Yaskawa INFORM job: KANT1.JBI

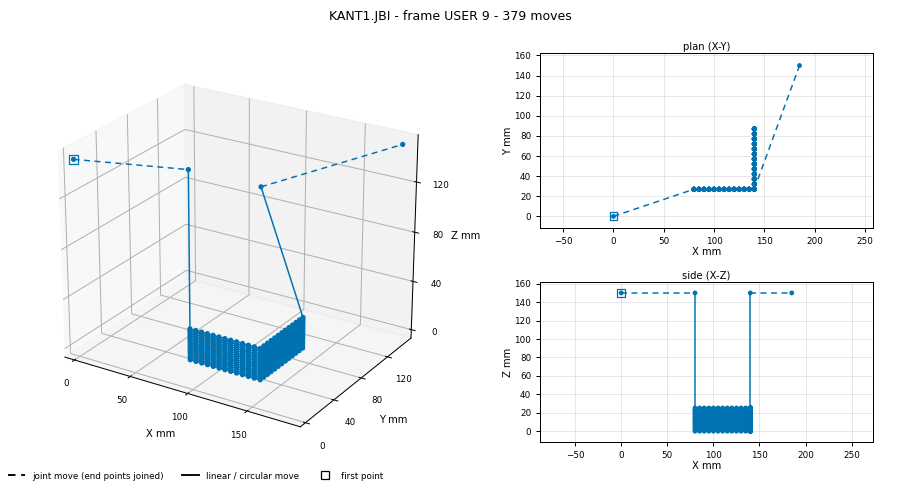
[picture p0: tool path of KANT1.JBI in frame USER 9, 379 of 379 moves have a stored position in this frame; points joined in program order, loops and branches not executed]
/JOB
//NAME KANT1
//POS
///NPOS 379,0,0,0,0,0
///USER 9
///TOOL 1
///POSTYPE USER
///RECTAN
///RCONF 1,0,0,0,0,0,0,0,0,0,0,0,0,0,0,0,0,0,0,0,0,0,0,0
C00000=0.000,0.000,150.000,0.0000,0.0000,-170.0000
C00001=80.000,27.000,150.000,0.0000,0.0000,-170.0000
C00002=80.000,27.000,0.000,0.0000,0.0000,-170.0000
C00003=85.000,27.000,0.000,0.0000,0.0000,-170.0000
C00004=90.000,27.000,0.000,0.0000,0.0000,-170.0000
C00005=95.000,27.000,0.000,0.0000,0.0000,-170.0000
C00006=100.000,27.000,0.000,0.0000,0.0000,-170.0000
C00007=105.000,27.000,0.000,0.0000,0.0000,-170.0000
C00008=110.000,27.000,0.000,0.0000,0.0000,-170.0000
C00009=115.000,27.000,0.000,0.0000,0.0000,-170.0000
C00010=120.000,27.000,0.000,0.0000,0.0000,-170.0000
C00011=125.000,27.000,0.000,0.0000,0.0000,-170.0000
C00012=130.000,27.000,0.000,0.0000,0.0000,-170.0000
C00013=135.000,27.000,0.000,0.0000,0.0000,-170.0000
C00014=140.000,27.000,0.000,0.0000,0.0000,-170.0000
C00015=140.000,32.000,0.000,0.0000,0.0000,-170.0000
C00016=140.000,37.000,0.000,0.0000,0.0000,-170.0000
C00017=140.000,42.000,0.000,0.0000,0.0000,-170.0000
C00018=140.000,47.000,0.000,0.0000,0.0000,-170.0000
C00019=140.000,52.000,0.000,0.0000,0.0000,-170.0000
C00020=140.000,57.000,0.000,0.0000,0.0000,-170.0000
C00021=140.000,62.000,0.000,0.0000,0.0000,-170.0000
C00022=140.000,67.000,0.000,0.0000,0.0000,-170.0000
C00023=140.000,72.000,0.000,0.0000,0.0000,-170.0000
C00024=140.000,77.000,0.000,0.0000,0.0000,-170.0000
C00025=140.000,82.000,0.000,0.0000,0.0000,-170.0000
C00026=140.000,87.000,0.000,0.0000,0.0000,-170.0000
C00027=140.000,87.000,1.800,0.0000,0.0000,-170.0000
C00028=140.000,82.000,1.800,0.0000,0.0000,-170.0000
C00029=140.000,77.000,1.800,0.0000,0.0000,-170.0000
C00030=140.000,72.000,1.800,0.0000,0.0000,-170.0000
C00031=140.000,67.000,1.800,0.0000,0.0000,-170.0000
C00032=140.000,62.000,1.800,0.0000,0.0000,-170.0000
C00033=140.000,57.000,1.800,0.0000,0.0000,-170.0000
C00034=140.000,52.000,1.800,0.0000,0.0000,-170.0000
C00035=140.000,47.000,1.800,0.0000,0.0000,-170.0000
C00036=140.000,42.000,1.800,0.0000,0.0000,-170.0000
C00037=140.000,37.000,1.800,0.0000,0.0000,-170.0000
C00038=140.000,32.000,1.800,0.0000,0.0000,-170.0000
C00039=140.000,27.000,1.800,0.0000,0.0000,-170.0000
C00040=135.000,27.000,1.800,0.0000,0.0000,-170.0000
C00041=130.000,27.000,1.800,0.0000,0.0000,-170.0000
C00042=125.000,27.000,1.800,0.0000,0.0000,-170.0000
C00043=120.000,27.000,1.800,0.0000,0.0000,-170.0000
C00044=115.000,27.000,1.800,0.0000,0.0000,-170.0000
C00045=110.000,27.000,1.800,0.0000,0.0000,-170.0000
C00046=105.000,27.000,1.800,0.0000,0.0000,-170.0000
C00047=100.000,27.000,1.800,0.0000,0.0000,-170.0000
C00048=95.000,27.000,1.800,0.0000,0.0000,-170.0000
C00049=90.000,27.000,1.800,0.0000,0.0000,-170.0000
C00050=85.000,27.000,1.800,0.0000,0.0000,-170.0000
C00051=80.000,27.000,1.800,0.0000,0.0000,-170.0000
C00052=80.000,27.000,3.600,0.0000,0.0000,-170.0000
C00053=85.000,27.000,3.600,0.0000,0.0000,-170.0000
C00054=90.000,27.000,3.600,0.0000,0.0000,-170.0000
C00055=95.000,27.000,3.600,0.0000,0.0000,-170.0000
C00056=100.000,27.000,3.600,0.0000,0.0000,-170.0000
C00057=105.000,27.000,3.600,0.0000,0.0000,-170.0000
C00058=110.000,27.000,3.600,0.0000,0.0000,-170.0000
C00059=115.000,27.000,3.600,0.0000,0.0000,-170.0000
C00060=120.000,27.000,3.600,0.0000,0.0000,-170.0000
C00061=125.000,27.000,3.600,0.0000,0.0000,-170.0000
C00062=130.000,27.000,3.600,0.0000,0.0000,-170.0000
C00063=135.000,27.000,3.600,0.0000,0.0000,-170.0000
C00064=140.000,27.000,3.600,0.0000,0.0000,-170.0000
C00065=140.000,32.000,3.600,0.0000,0.0000,-170.0000
C00066=140.000,37.000,3.600,0.0000,0.0000,-170.0000
C00067=140.000,42.000,3.600,0.0000,0.0000,-170.0000
C00068=140.000,47.000,3.600,0.0000,0.0000,-170.0000
C00069=140.000,52.000,3.600,0.0000,0.0000,-170.0000
C00070=140.000,57.000,3.600,0.0000,0.0000,-170.0000
C00071=140.000,62.000,3.600,0.0000,0.0000,-170.0000
C00072=140.000,67.000,3.600,0.0000,0.0000,-170.0000
C00073=140.000,72.000,3.600,0.0000,0.0000,-170.0000
C00074=140.000,77.000,3.600,0.0000,0.0000,-170.0000
C00075=140.000,82.000,3.600,0.0000,0.0000,-170.0000
C00076=140.000,87.000,3.600,0.0000,0.0000,-170.0000
C00077=140.000,87.000,5.400,0.0000,0.0000,-170.0000
C00078=140.000,82.000,5.400,0.0000,0.0000,-170.0000
C00079=140.000,77.000,5.400,0.0000,0.0000,-170.0000
C00080=140.000,72.000,5.400,0.0000,0.0000,-170.0000
C00081=140.000,67.000,5.400,0.0000,0.0000,-170.0000
C00082=140.000,62.000,5.400,0.0000,0.0000,-170.0000
C00083=140.000,57.000,5.400,0.0000,0.0000,-170.0000
C00084=140.000,52.000,5.400,0.0000,0.0000,-170.0000
C00085=140.000,47.000,5.400,0.0000,0.0000,-170.0000
C00086=140.000,42.000,5.400,0.0000,0.0000,-170.0000
C00087=140.000,37.000,5.400,0.0000,0.0000,-170.0000
C00088=140.000,32.000,5.400,0.0000,0.0000,-170.0000
C00089=140.000,27.000,5.400,0.0000,0.0000,-170.0000
C00090=135.000,27.000,5.400,0.0000,0.0000,-170.0000
C00091=130.000,27.000,5.400,0.0000,0.0000,-170.0000
C00092=125.000,27.000,5.400,0.0000,0.0000,-170.0000
C00093=120.000,27.000,5.400,0.0000,0.0000,-170.0000
C00094=115.000,27.000,5.400,0.0000,0.0000,-170.0000
C00095=110.000,27.000,5.400,0.0000,0.0000,-170.0000
C00096=105.000,27.000,5.400,0.0000,0.0000,-170.0000
C00097=100.000,27.000,5.400,0.0000,0.0000,-170.0000
C00098=95.000,27.000,5.400,0.0000,0.0000,-170.0000
C00099=90.000,27.000,5.400,0.0000,0.0000,-170.0000
C00100=85.000,27.000,5.400,0.0000,0.0000,-170.0000
C00101=80.000,27.000,5.400,0.0000,0.0000,-170.0000
C00102=80.000,27.000,7.200,0.0000,0.0000,-170.0000
C00103=85.000,27.000,7.200,0.0000,0.0000,-170.0000
C00104=90.000,27.000,7.200,0.0000,0.0000,-170.0000
C00105=95.000,27.000,7.200,0.0000,0.0000,-170.0000
C00106=100.000,27.000,7.200,0.0000,0.0000,-170.0000
C00107=105.000,27.000,7.200,0.0000,0.0000,-170.0000
C00108=110.000,27.000,7.200,0.0000,0.0000,-170.0000
C00109=115.000,27.000,7.200,0.0000,0.0000,-170.0000
C00110=120.000,27.000,7.200,0.0000,0.0000,-170.0000
C00111=125.000,27.000,7.200,0.0000,0.0000,-170.0000
C00112=130.000,27.000,7.200,0.0000,0.0000,-170.0000
C00113=135.000,27.000,7.200,0.0000,0.0000,-170.0000
C00114=140.000,27.000,7.200,0.0000,0.0000,-170.0000
C00115=140.000,32.000,7.200,0.0000,0.0000,-170.0000
C00116=140.000,37.000,7.200,0.0000,0.0000,-170.0000
C00117=140.000,42.000,7.200,0.0000,0.0000,-170.0000
C00118=140.000,47.000,7.200,0.0000,0.0000,-170.0000
C00119=140.000,52.000,7.200,0.0000,0.0000,-170.0000
C00120=140.000,57.000,7.200,0.0000,0.0000,-170.0000
C00121=140.000,62.000,7.200,0.0000,0.0000,-170.0000
C00122=140.000,67.000,7.200,0.0000,0.0000,-170.0000
C00123=140.000,72.000,7.200,0.0000,0.0000,-170.0000
C00124=140.000,77.000,7.200,0.0000,0.0000,-170.0000
C00125=140.000,82.000,7.200,0.0000,0.0000,-170.0000
C00126=140.000,87.000,7.200,0.0000,0.0000,-170.0000
C00127=140.000,87.000,9.000,0.0000,0.0000,-170.0000
C00128=140.000,82.000,9.000,0.0000,0.0000,-170.0000
C00129=140.000,77.000,9.000,0.0000,0.0000,-170.0000
C00130=140.000,72.000,9.000,0.0000,0.0000,-170.0000
C00131=140.000,67.000,9.000,0.0000,0.0000,-170.0000
C00132=140.000,62.000,9.000,0.0000,0.0000,-170.0000
C00133=140.000,57.000,9.000,0.0000,0.0000,-170.0000
C00134=140.000,52.000,9.000,0.0000,0.0000,-170.0000
C00135=140.000,47.000,9.000,0.0000,0.0000,-170.0000
C00136=140.000,42.000,9.000,0.0000,0.0000,-170.0000
C00137=140.000,37.000,9.000,0.0000,0.0000,-170.0000
C00138=140.000,32.000,9.000,0.0000,0.0000,-170.0000
C00139=140.000,27.000,9.000,0.0000,0.0000,-170.0000
C00140=135.000,27.000,9.000,0.0000,0.0000,-170.0000
C00141=130.000,27.000,9.000,0.0000,0.0000,-170.0000
C00142=125.000,27.000,9.000,0.0000,0.0000,-170.0000
C00143=120.000,27.000,9.000,0.0000,0.0000,-170.0000
C00144=115.000,27.000,9.000,0.0000,0.0000,-170.0000
C00145=110.000,27.000,9.000,0.0000,0.0000,-170.0000
C00146=105.000,27.000,9.000,0.0000,0.0000,-170.0000
C00147=100.000,27.000,9.000,0.0000,0.0000,-170.0000
C00148=95.000,27.000,9.000,0.0000,0.0000,-170.0000
C00149=90.000,27.000,9.000,0.0000,0.0000,-170.0000
C00150=85.000,27.000,9.000,0.0000,0.0000,-170.0000
C00151=80.000,27.000,9.000,0.0000,0.0000,-170.0000
C00152=80.000,27.000,10.800,0.0000,0.0000,-170.0000
C00153=85.000,27.000,10.800,0.0000,0.0000,-170.0000
C00154=90.000,27.000,10.800,0.0000,0.0000,-170.0000
C00155=95.000,27.000,10.800,0.0000,0.0000,-170.0000
C00156=100.000,27.000,10.800,0.0000,0.0000,-170.0000
C00157=105.000,27.000,10.800,0.0000,0.0000,-170.0000
C00158=110.000,27.000,10.800,0.0000,0.0000,-170.0000
C00159=115.000,27.000,10.800,0.0000,0.0000,-170.0000
C00160=120.000,27.000,10.800,0.0000,0.0000,-170.0000
C00161=125.000,27.000,10.800,0.0000,0.0000,-170.0000
C00162=130.000,27.000,10.800,0.0000,0.0000,-170.0000
C00163=135.000,27.000,10.800,0.0000,0.0000,-170.0000
C00164=140.000,27.000,10.800,0.0000,0.0000,-170.0000
C00165=140.000,32.000,10.800,0.0000,0.0000,-170.0000
C00166=140.000,37.000,10.800,0.0000,0.0000,-170.0000
C00167=140.000,42.000,10.800,0.0000,0.0000,-170.0000
C00168=140.000,47.000,10.800,0.0000,0.0000,-170.0000
C00169=140.000,52.000,10.800,0.0000,0.0000,-170.0000
C00170=140.000,57.000,10.800,0.0000,0.0000,-170.0000
C00171=140.000,62.000,10.800,0.0000,0.0000,-170.0000
C00172=140.000,67.000,10.800,0.0000,0.0000,-170.0000
C00173=140.000,72.000,10.800,0.0000,0.0000,-170.0000
C00174=140.000,77.000,10.800,0.0000,0.0000,-170.0000
C00175=140.000,82.000,10.800,0.0000,0.0000,-170.0000
C00176=140.000,87.000,10.800,0.0000,0.0000,-170.0000
C00177=140.000,87.000,12.600,0.0000,0.0000,-170.0000
C00178=140.000,82.000,12.600,0.0000,0.0000,-170.0000
C00179=140.000,77.000,12.600,0.0000,0.0000,-170.0000
C00180=140.000,72.000,12.600,0.0000,0.0000,-170.0000
C00181=140.000,67.000,12.600,0.0000,0.0000,-170.0000
C00182=140.000,62.000,12.600,0.0000,0.0000,-170.0000
C00183=140.000,57.000,12.600,0.0000,0.0000,-170.0000
C00184=140.000,52.000,12.600,0.0000,0.0000,-170.0000
C00185=140.000,47.000,12.600,0.0000,0.0000,-170.0000
C00186=140.000,42.000,12.600,0.0000,0.0000,-170.0000
C00187=140.000,37.000,12.600,0.0000,0.0000,-170.0000
C00188=140.000,32.000,12.600,0.0000,0.0000,-170.0000
C00189=140.000,27.000,12.600,0.0000,0.0000,-170.0000
C00190=135.000,27.000,12.600,0.0000,0.0000,-170.0000
C00191=130.000,27.000,12.600,0.0000,0.0000,-170.0000
C00192=125.000,27.000,12.600,0.0000,0.0000,-170.0000
C00193=120.000,27.000,12.600,0.0000,0.0000,-170.0000
C00194=115.000,27.000,12.600,0.0000,0.0000,-170.0000
C00195=110.000,27.000,12.600,0.0000,0.0000,-170.0000
C00196=105.000,27.000,12.600,0.0000,0.0000,-170.0000
C00197=100.000,27.000,12.600,0.0000,0.0000,-170.0000
C00198=95.000,27.000,12.600,0.0000,0.0000,-170.0000
C00199=90.000,27.000,12.600,0.0000,0.0000,-170.0000
C00200=85.000,27.000,12.600,0.0000,0.0000,-170.0000
C00201=80.000,27.000,12.600,0.0000,0.0000,-170.0000
C00202=80.000,27.000,14.400,0.0000,0.0000,-170.0000
C00203=85.000,27.000,14.400,0.0000,0.0000,-170.0000
C00204=90.000,27.000,14.400,0.0000,0.0000,-170.0000
C00205=95.000,27.000,14.400,0.0000,0.0000,-170.0000
C00206=100.000,27.000,14.400,0.0000,0.0000,-170.0000
C00207=105.000,27.000,14.400,0.0000,0.0000,-170.0000
C00208=110.000,27.000,14.400,0.0000,0.0000,-170.0000
C00209=115.000,27.000,14.400,0.0000,0.0000,-170.0000
C00210=120.000,27.000,14.400,0.0000,0.0000,-170.0000
C00211=125.000,27.000,14.400,0.0000,0.0000,-170.0000
C00212=130.000,27.000,14.400,0.0000,0.0000,-170.0000
C00213=135.000,27.000,14.400,0.0000,0.0000,-170.0000
C00214=140.000,27.000,14.400,0.0000,0.0000,-170.0000
C00215=140.000,32.000,14.400,0.0000,0.0000,-170.0000
C00216=140.000,37.000,14.400,0.0000,0.0000,-170.0000
C00217=140.000,42.000,14.400,0.0000,0.0000,-170.0000
C00218=140.000,47.000,14.400,0.0000,0.0000,-170.0000
C00219=140.000,52.000,14.400,0.0000,0.0000,-170.0000
C00220=140.000,57.000,14.400,0.0000,0.0000,-170.0000
C00221=140.000,62.000,14.400,0.0000,0.0000,-170.0000
C00222=140.000,67.000,14.400,0.0000,0.0000,-170.0000
C00223=140.000,72.000,14.400,0.0000,0.0000,-170.0000
C00224=140.000,77.000,14.400,0.0000,0.0000,-170.0000
C00225=140.000,82.000,14.400,0.0000,0.0000,-170.0000
C00226=140.000,87.000,14.400,0.0000,0.0000,-170.0000
C00227=140.000,87.000,16.200,0.0000,0.0000,-170.0000
C00228=140.000,82.000,16.200,0.0000,0.0000,-170.0000
C00229=140.000,77.000,16.200,0.0000,0.0000,-170.0000
C00230=140.000,72.000,16.200,0.0000,0.0000,-170.0000
C00231=140.000,67.000,16.200,0.0000,0.0000,-170.0000
C00232=140.000,62.000,16.200,0.0000,0.0000,-170.0000
C00233=140.000,57.000,16.200,0.0000,0.0000,-170.0000
C00234=140.000,52.000,16.200,0.0000,0.0000,-170.0000
C00235=140.000,47.000,16.200,0.0000,0.0000,-170.0000
C00236=140.000,42.000,16.200,0.0000,0.0000,-170.0000
C00237=140.000,37.000,16.200,0.0000,0.0000,-170.0000
C00238=140.000,32.000,16.200,0.0000,0.0000,-170.0000
C00239=140.000,27.000,16.200,0.0000,0.0000,-170.0000
C00240=135.000,27.000,16.200,0.0000,0.0000,-170.0000
C00241=130.000,27.000,16.200,0.0000,0.0000,-170.0000
C00242=125.000,27.000,16.200,0.0000,0.0000,-170.0000
C00243=120.000,27.000,16.200,0.0000,0.0000,-170.0000
C00244=115.000,27.000,16.200,0.0000,0.0000,-170.0000
C00245=110.000,27.000,16.200,0.0000,0.0000,-170.0000
C00246=105.000,27.000,16.200,0.0000,0.0000,-170.0000
C00247=100.000,27.000,16.200,0.0000,0.0000,-170.0000
C00248=95.000,27.000,16.200,0.0000,0.0000,-170.0000
C00249=90.000,27.000,16.200,0.0000,0.0000,-170.0000
C00250=85.000,27.000,16.200,0.0000,0.0000,-170.0000
C00251=80.000,27.000,16.200,0.0000,0.0000,-170.0000
C00252=80.000,27.000,18.000,0.0000,0.0000,-170.0000
C00253=85.000,27.000,18.000,0.0000,0.0000,-170.0000
C00254=90.000,27.000,18.000,0.0000,0.0000,-170.0000
C00255=95.000,27.000,18.000,0.0000,0.0000,-170.0000
C00256=100.000,27.000,18.000,0.0000,0.0000,-170.0000
C00257=105.000,27.000,18.000,0.0000,0.0000,-170.0000
C00258=110.000,27.000,18.000,0.0000,0.0000,-170.0000
C00259=115.000,27.000,18.000,0.0000,0.0000,-170.0000
C00260=120.000,27.000,18.000,0.0000,0.0000,-170.0000
C00261=125.000,27.000,18.000,0.0000,0.0000,-170.0000
C00262=130.000,27.000,18.000,0.0000,0.0000,-170.0000
C00263=135.000,27.000,18.000,0.0000,0.0000,-170.0000
C00264=140.000,27.000,18.000,0.0000,0.0000,-170.0000
C00265=140.000,32.000,18.000,0.0000,0.0000,-170.0000
C00266=140.000,37.000,18.000,0.0000,0.0000,-170.0000
C00267=140.000,42.000,18.000,0.0000,0.0000,-170.0000
C00268=140.000,47.000,18.000,0.0000,0.0000,-170.0000
C00269=140.000,52.000,18.000,0.0000,0.0000,-170.0000
C00270=140.000,57.000,18.000,0.0000,0.0000,-170.0000
C00271=140.000,62.000,18.000,0.0000,0.0000,-170.0000
C00272=140.000,67.000,18.000,0.0000,0.0000,-170.0000
C00273=140.000,72.000,18.000,0.0000,0.0000,-170.0000
C00274=140.000,77.000,18.000,0.0000,0.0000,-170.0000
C00275=140.000,82.000,18.000,0.0000,0.0000,-170.0000
C00276=140.000,87.000,18.000,0.0000,0.0000,-170.0000
C00277=140.000,87.000,19.800,0.0000,0.0000,-170.0000
C00278=140.000,82.000,19.800,0.0000,0.0000,-170.0000
C00279=140.000,77.000,19.800,0.0000,0.0000,-170.0000
C00280=140.000,72.000,19.800,0.0000,0.0000,-170.0000
C00281=140.000,67.000,19.800,0.0000,0.0000,-170.0000
C00282=140.000,62.000,19.800,0.0000,0.0000,-170.0000
C00283=140.000,57.000,19.800,0.0000,0.0000,-170.0000
C00284=140.000,52.000,19.800,0.0000,0.0000,-170.0000
C00285=140.000,47.000,19.800,0.0000,0.0000,-170.0000
C00286=140.000,42.000,19.800,0.0000,0.0000,-170.0000
C00287=140.000,37.000,19.800,0.0000,0.0000,-170.0000
C00288=140.000,32.000,19.800,0.0000,0.0000,-170.0000
C00289=140.000,27.000,19.800,0.0000,0.0000,-170.0000
C00290=135.000,27.000,19.800,0.0000,0.0000,-170.0000
C00291=130.000,27.000,19.800,0.0000,0.0000,-170.0000
C00292=125.000,27.000,19.800,0.0000,0.0000,-170.0000
C00293=120.000,27.000,19.800,0.0000,0.0000,-170.0000
C00294=115.000,27.000,19.800,0.0000,0.0000,-170.0000
C00295=110.000,27.000,19.800,0.0000,0.0000,-170.0000
C00296=105.000,27.000,19.800,0.0000,0.0000,-170.0000
C00297=100.000,27.000,19.800,0.0000,0.0000,-170.0000
C00298=95.000,27.000,19.800,0.0000,0.0000,-170.0000
C00299=90.000,27.000,19.800,0.0000,0.0000,-170.0000
C00300=85.000,27.000,19.800,0.0000,0.0000,-170.0000
C00301=80.000,27.000,19.800,0.0000,0.0000,-170.0000
C00302=80.000,27.000,21.600,0.0000,0.0000,-170.0000
C00303=85.000,27.000,21.600,0.0000,0.0000,-170.0000
C00304=90.000,27.000,21.600,0.0000,0.0000,-170.0000
C00305=95.000,27.000,21.600,0.0000,0.0000,-170.0000
C00306=100.000,27.000,21.600,0.0000,0.0000,-170.0000
C00307=105.000,27.000,21.600,0.0000,0.0000,-170.0000
C00308=110.000,27.000,21.600,0.0000,0.0000,-170.0000
C00309=115.000,27.000,21.600,0.0000,0.0000,-170.0000
C00310=120.000,27.000,21.600,0.0000,0.0000,-170.0000
C00311=125.000,27.000,21.600,0.0000,0.0000,-170.0000
C00312=130.000,27.000,21.600,0.0000,0.0000,-170.0000
C00313=135.000,27.000,21.600,0.0000,0.0000,-170.0000
C00314=140.000,27.000,21.600,0.0000,0.0000,-170.0000
C00315=140.000,32.000,21.600,0.0000,0.0000,-170.0000
C00316=140.000,37.000,21.600,0.0000,0.0000,-170.0000
C00317=140.000,42.000,21.600,0.0000,0.0000,-170.0000
C00318=140.000,47.000,21.600,0.0000,0.0000,-170.0000
C00319=140.000,52.000,21.600,0.0000,0.0000,-170.0000
C00320=140.000,57.000,21.600,0.0000,0.0000,-170.0000
C00321=140.000,62.000,21.600,0.0000,0.0000,-170.0000
C00322=140.000,67.000,21.600,0.0000,0.0000,-170.0000
C00323=140.000,72.000,21.600,0.0000,0.0000,-170.0000
C00324=140.000,77.000,21.600,0.0000,0.0000,-170.0000
C00325=140.000,82.000,21.600,0.0000,0.0000,-170.0000
C00326=140.000,87.000,21.600,0.0000,0.0000,-170.0000
C00327=140.000,87.000,23.400,0.0000,0.0000,-170.0000
C00328=140.000,82.000,23.400,0.0000,0.0000,-170.0000
C00329=140.000,77.000,23.400,0.0000,0.0000,-170.0000
C00330=140.000,72.000,23.400,0.0000,0.0000,-170.0000
C00331=140.000,67.000,23.400,0.0000,0.0000,-170.0000
C00332=140.000,62.000,23.400,0.0000,0.0000,-170.0000
C00333=140.000,57.000,23.400,0.0000,0.0000,-170.0000
C00334=140.000,52.000,23.400,0.0000,0.0000,-170.0000
C00335=140.000,47.000,23.400,0.0000,0.0000,-170.0000
C00336=140.000,42.000,23.400,0.0000,0.0000,-170.0000
C00337=140.000,37.000,23.400,0.0000,0.0000,-170.0000
C00338=140.000,32.000,23.400,0.0000,0.0000,-170.0000
C00339=140.000,27.000,23.400,0.0000,0.0000,-170.0000
C00340=135.000,27.000,23.400,0.0000,0.0000,-170.0000
C00341=130.000,27.000,23.400,0.0000,0.0000,-170.0000
C00342=125.000,27.000,23.400,0.0000,0.0000,-170.0000
C00343=120.000,27.000,23.400,0.0000,0.0000,-170.0000
C00344=115.000,27.000,23.400,0.0000,0.0000,-170.0000
C00345=110.000,27.000,23.400,0.0000,0.0000,-170.0000
C00346=105.000,27.000,23.400,0.0000,0.0000,-170.0000
C00347=100.000,27.000,23.400,0.0000,0.0000,-170.0000
C00348=95.000,27.000,23.400,0.0000,0.0000,-170.0000
C00349=90.000,27.000,23.400,0.0000,0.0000,-170.0000
C00350=85.000,27.000,23.400,0.0000,0.0000,-170.0000
C00351=80.000,27.000,23.400,0.0000,0.0000,-170.0000
C00352=80.000,27.000,25.200,0.0000,0.0000,-170.0000
C00353=85.000,27.000,25.200,0.0000,0.0000,-170.0000
C00354=90.000,27.000,25.200,0.0000,0.0000,-170.0000
C00355=95.000,27.000,25.200,0.0000,0.0000,-170.0000
C00356=100.000,27.000,25.200,0.0000,0.0000,-170.0000
C00357=105.000,27.000,25.200,0.0000,0.0000,-170.0000
C00358=110.000,27.000,25.200,0.0000,0.0000,-170.0000
C00359=115.000,27.000,25.200,0.0000,0.0000,-170.0000
C00360=120.000,27.000,25.200,0.0000,0.0000,-170.0000
C00361=125.000,27.000,25.200,0.0000,0.0000,-170.0000
C00362=130.000,27.000,25.200,0.0000,0.0000,-170.0000
C00363=135.000,27.000,25.200,0.0000,0.0000,-170.0000
C00364=140.000,27.000,25.200,0.0000,0.0000,-170.0000
C00365=140.000,32.000,25.200,0.0000,0.0000,-170.0000
C00366=140.000,37.000,25.200,0.0000,0.0000,-170.0000
C00367=140.000,42.000,25.200,0.0000,0.0000,-170.0000
C00368=140.000,47.000,25.200,0.0000,0.0000,-170.0000
C00369=140.000,52.000,25.200,0.0000,0.0000,-170.0000
C00370=140.000,57.000,25.200,0.0000,0.0000,-170.0000
C00371=140.000,62.000,25.200,0.0000,0.0000,-170.0000
C00372=140.000,67.000,25.200,0.0000,0.0000,-170.0000
C00373=140.000,72.000,25.200,0.0000,0.0000,-170.0000
C00374=140.000,77.000,25.200,0.0000,0.0000,-170.0000
C00375=140.000,82.000,25.200,0.0000,0.0000,-170.0000
C00376=140.000,87.000,25.200,0.0000,0.0000,-170.0000
C00377=140.000,27.000,150.000,0.0000,0.0000,-170.0000
C00378=185.000,150.000,150.000,0.0000,0.0000,-170.0000
//INST
///DATE 2026/10/23 16:08
///ATTR SC,RW,RJ
////FRAME USER 9
///GROUP1 RB1
NOP
MOVJ C00000 VJ=0.78
MOVJ C00001 VJ=0.78
MOVL C00002 V=11.0 ACC=20 DEC=20
*LAG1
MACRO1 MJ#(0) ARGF1
ARCON
MOVL C00003 V=7.0 ACC=20 DEC=20
MOVL C00004 V=7.0 ACC=20 DEC=20
MOVL C00005 V=7.0 ACC=20 DEC=20
MOVL C00006 V=7.0 ACC=20 DEC=20
MOVL C00007 V=7.0 ACC=20 DEC=20
MOVL C00008 V=7.0 ACC=20 DEC=20
MOVL C00009 V=7.0 ACC=20 DEC=20
MOVL C00010 V=7.0 ACC=20 DEC=20
MOVL C00011 V=7.0 ACC=20 DEC=20
MOVL C00012 V=7.0 ACC=20 DEC=20
MOVL C00013 V=7.0 ACC=20 DEC=20
MOVL C00014 V=7.0 ACC=20 DEC=20
MOVL C00015 V=7.0 ACC=20 DEC=20
MOVL C00016 V=7.0 ACC=20 DEC=20
MOVL C00017 V=7.0 ACC=20 DEC=20
MOVL C00018 V=7.0 ACC=20 DEC=20
MOVL C00019 V=7.0 ACC=20 DEC=20
MOVL C00020 V=7.0 ACC=20 DEC=20
MOVL C00021 V=7.0 ACC=20 DEC=20
MOVL C00022 V=7.0 ACC=20 DEC=20
MOVL C00023 V=7.0 ACC=20 DEC=20
MOVL C00024 V=7.0 ACC=20 DEC=20
MOVL C00025 V=7.0 ACC=20 DEC=20
MOVL C00026 V=7.0 ACC=20 DEC=20
ARCOF
TIMER T=30
*LAG2
MOVL C00027 V=11.0 ACC=20 DEC=20
MACRO1 MJ#(0) ARGF2
ARCON
MOVL C00028 V=7.0 ACC=20 DEC=20
MOVL C00029 V=7.0 ACC=20 DEC=20
MOVL C00030 V=7.0 ACC=20 DEC=20
MOVL C00031 V=7.0 ACC=20 DEC=20
MOVL C00032 V=7.0 ACC=20 DEC=20
MOVL C00033 V=7.0 ACC=20 DEC=20
MOVL C00034 V=7.0 ACC=20 DEC=20
MOVL C00035 V=7.0 ACC=20 DEC=20
MOVL C00036 V=7.0 ACC=20 DEC=20
MOVL C00037 V=7.0 ACC=20 DEC=20
MOVL C00038 V=7.0 ACC=20 DEC=20
MOVL C00039 V=7.0 ACC=20 DEC=20
MOVL C00040 V=7.0 ACC=20 DEC=20
MOVL C00041 V=7.0 ACC=20 DEC=20
MOVL C00042 V=7.0 ACC=20 DEC=20
MOVL C00043 V=7.0 ACC=20 DEC=20
MOVL C00044 V=7.0 ACC=20 DEC=20
MOVL C00045 V=7.0 ACC=20 DEC=20
MOVL C00046 V=7.0 ACC=20 DEC=20
MOVL C00047 V=7.0 ACC=20 DEC=20
MOVL C00048 V=7.0 ACC=20 DEC=20
MOVL C00049 V=7.0 ACC=20 DEC=20
MOVL C00050 V=7.0 ACC=20 DEC=20
MOVL C00051 V=7.0 ACC=20 DEC=20
ARCOF
TIMER T=30
*LAG3
MOVL C00052 V=11.0 ACC=20 DEC=20
MACRO1 MJ#(0) ARGF2
ARCON
MOVL C00053 V=7.0 ACC=20 DEC=20
MOVL C00054 V=7.0 ACC=20 DEC=20
MOVL C00055 V=7.0 ACC=20 DEC=20
MOVL C00056 V=7.0 ACC=20 DEC=20
MOVL C00057 V=7.0 ACC=20 DEC=20
MOVL C00058 V=7.0 ACC=20 DEC=20
MOVL C00059 V=7.0 ACC=20 DEC=20
MOVL C00060 V=7.0 ACC=20 DEC=20
MOVL C00061 V=7.0 ACC=20 DEC=20
MOVL C00062 V=7.0 ACC=20 DEC=20
MOVL C00063 V=7.0 ACC=20 DEC=20
MOVL C00064 V=7.0 ACC=20 DEC=20
MOVL C00065 V=7.0 ACC=20 DEC=20
MOVL C00066 V=7.0 ACC=20 DEC=20
MOVL C00067 V=7.0 ACC=20 DEC=20
MOVL C00068 V=7.0 ACC=20 DEC=20
MOVL C00069 V=7.0 ACC=20 DEC=20
MOVL C00070 V=7.0 ACC=20 DEC=20
MOVL C00071 V=7.0 ACC=20 DEC=20
MOVL C00072 V=7.0 ACC=20 DEC=20
MOVL C00073 V=7.0 ACC=20 DEC=20
MOVL C00074 V=7.0 ACC=20 DEC=20
MOVL C00075 V=7.0 ACC=20 DEC=20
MOVL C00076 V=7.0 ACC=20 DEC=20
ARCOF
TIMER T=30
*LAG4
MOVL C00077 V=11.0 ACC=20 DEC=20
MACRO1 MJ#(0) ARGF2
ARCON
MOVL C00078 V=7.0 ACC=20 DEC=20
MOVL C00079 V=7.0 ACC=20 DEC=20
MOVL C00080 V=7.0 ACC=20 DEC=20
MOVL C00081 V=7.0 ACC=20 DEC=20
MOVL C00082 V=7.0 ACC=20 DEC=20
MOVL C00083 V=7.0 ACC=20 DEC=20
MOVL C00084 V=7.0 ACC=20 DEC=20
MOVL C00085 V=7.0 ACC=20 DEC=20
MOVL C00086 V=7.0 ACC=20 DEC=20
MOVL C00087 V=7.0 ACC=20 DEC=20
MOVL C00088 V=7.0 ACC=20 DEC=20
MOVL C00089 V=7.0 ACC=20 DEC=20
MOVL C00090 V=7.0 ACC=20 DEC=20
MOVL C00091 V=7.0 ACC=20 DEC=20
MOVL C00092 V=7.0 ACC=20 DEC=20
MOVL C00093 V=7.0 ACC=20 DEC=20
MOVL C00094 V=7.0 ACC=20 DEC=20
MOVL C00095 V=7.0 ACC=20 DEC=20
MOVL C00096 V=7.0 ACC=20 DEC=20
MOVL C00097 V=7.0 ACC=20 DEC=20
MOVL C00098 V=7.0 ACC=20 DEC=20
MOVL C00099 V=7.0 ACC=20 DEC=20
MOVL C00100 V=7.0 ACC=20 DEC=20
MOVL C00101 V=7.0 ACC=20 DEC=20
ARCOF
TIMER T=30
*LAG5
MOVL C00102 V=11.0 ACC=20 DEC=20
MACRO1 MJ#(0) ARGF2
ARCON
MOVL C00103 V=7.0 ACC=20 DEC=20
MOVL C00104 V=7.0 ACC=20 DEC=20
MOVL C00105 V=7.0 ACC=20 DEC=20
MOVL C00106 V=7.0 ACC=20 DEC=20
MOVL C00107 V=7.0 ACC=20 DEC=20
MOVL C00108 V=7.0 ACC=20 DEC=20
MOVL C00109 V=7.0 ACC=20 DEC=20
MOVL C00110 V=7.0 ACC=20 DEC=20
MOVL C00111 V=7.0 ACC=20 DEC=20
MOVL C00112 V=7.0 ACC=20 DEC=20
MOVL C00113 V=7.0 ACC=20 DEC=20
MOVL C00114 V=7.0 ACC=20 DEC=20
MOVL C00115 V=7.0 ACC=20 DEC=20
MOVL C00116 V=7.0 ACC=20 DEC=20
MOVL C00117 V=7.0 ACC=20 DEC=20
MOVL C00118 V=7.0 ACC=20 DEC=20
MOVL C00119 V=7.0 ACC=20 DEC=20
MOVL C00120 V=7.0 ACC=20 DEC=20
MOVL C00121 V=7.0 ACC=20 DEC=20
MOVL C00122 V=7.0 ACC=20 DEC=20
MOVL C00123 V=7.0 ACC=20 DEC=20
MOVL C00124 V=7.0 ACC=20 DEC=20
MOVL C00125 V=7.0 ACC=20 DEC=20
MOVL C00126 V=7.0 ACC=20 DEC=20
ARCOF
TIMER T=30
*LAG6
MOVL C00127 V=11.0 ACC=20 DEC=20
MACRO1 MJ#(0) ARGF2
ARCON
MOVL C00128 V=7.0 ACC=20 DEC=20
MOVL C00129 V=7.0 ACC=20 DEC=20
MOVL C00130 V=7.0 ACC=20 DEC=20
MOVL C00131 V=7.0 ACC=20 DEC=20
MOVL C00132 V=7.0 ACC=20 DEC=20
MOVL C00133 V=7.0 ACC=20 DEC=20
MOVL C00134 V=7.0 ACC=20 DEC=20
MOVL C00135 V=7.0 ACC=20 DEC=20
MOVL C00136 V=7.0 ACC=20 DEC=20
MOVL C00137 V=7.0 ACC=20 DEC=20
MOVL C00138 V=7.0 ACC=20 DEC=20
MOVL C00139 V=7.0 ACC=20 DEC=20
MOVL C00140 V=7.0 ACC=20 DEC=20
MOVL C00141 V=7.0 ACC=20 DEC=20
MOVL C00142 V=7.0 ACC=20 DEC=20
MOVL C00143 V=7.0 ACC=20 DEC=20
MOVL C00144 V=7.0 ACC=20 DEC=20
MOVL C00145 V=7.0 ACC=20 DEC=20
MOVL C00146 V=7.0 ACC=20 DEC=20
MOVL C00147 V=7.0 ACC=20 DEC=20
MOVL C00148 V=7.0 ACC=20 DEC=20
MOVL C00149 V=7.0 ACC=20 DEC=20
MOVL C00150 V=7.0 ACC=20 DEC=20
MOVL C00151 V=7.0 ACC=20 DEC=20
ARCOF
TIMER T=30
*LAG7
MOVL C00152 V=11.0 ACC=20 DEC=20
MACRO1 MJ#(0) ARGF2
ARCON
MOVL C00153 V=7.0 ACC=20 DEC=20
MOVL C00154 V=7.0 ACC=20 DEC=20
MOVL C00155 V=7.0 ACC=20 DEC=20
MOVL C00156 V=7.0 ACC=20 DEC=20
MOVL C00157 V=7.0 ACC=20 DEC=20
MOVL C00158 V=7.0 ACC=20 DEC=20
MOVL C00159 V=7.0 ACC=20 DEC=20
MOVL C00160 V=7.0 ACC=20 DEC=20
MOVL C00161 V=7.0 ACC=20 DEC=20
MOVL C00162 V=7.0 ACC=20 DEC=20
MOVL C00163 V=7.0 ACC=20 DEC=20
MOVL C00164 V=7.0 ACC=20 DEC=20
MOVL C00165 V=7.0 ACC=20 DEC=20
MOVL C00166 V=7.0 ACC=20 DEC=20
MOVL C00167 V=7.0 ACC=20 DEC=20
MOVL C00168 V=7.0 ACC=20 DEC=20
MOVL C00169 V=7.0 ACC=20 DEC=20
MOVL C00170 V=7.0 ACC=20 DEC=20
MOVL C00171 V=7.0 ACC=20 DEC=20
MOVL C00172 V=7.0 ACC=20 DEC=20
MOVL C00173 V=7.0 ACC=20 DEC=20
MOVL C00174 V=7.0 ACC=20 DEC=20
MOVL C00175 V=7.0 ACC=20 DEC=20
MOVL C00176 V=7.0 ACC=20 DEC=20
ARCOF
TIMER T=30
*LAG8
MOVL C00177 V=11.0 ACC=20 DEC=20
MACRO1 MJ#(0) ARGF2
ARCON
MOVL C00178 V=7.0 ACC=20 DEC=20
MOVL C00179 V=7.0 ACC=20 DEC=20
MOVL C00180 V=7.0 ACC=20 DEC=20
MOVL C00181 V=7.0 ACC=20 DEC=20
MOVL C00182 V=7.0 ACC=20 DEC=20
MOVL C00183 V=7.0 ACC=20 DEC=20
MOVL C00184 V=7.0 ACC=20 DEC=20
MOVL C00185 V=7.0 ACC=20 DEC=20
MOVL C00186 V=7.0 ACC=20 DEC=20
MOVL C00187 V=7.0 ACC=20 DEC=20
MOVL C00188 V=7.0 ACC=20 DEC=20
MOVL C00189 V=7.0 ACC=20 DEC=20
MOVL C00190 V=7.0 ACC=20 DEC=20
MOVL C00191 V=7.0 ACC=20 DEC=20
MOVL C00192 V=7.0 ACC=20 DEC=20
MOVL C00193 V=7.0 ACC=20 DEC=20
MOVL C00194 V=7.0 ACC=20 DEC=20
MOVL C00195 V=7.0 ACC=20 DEC=20
MOVL C00196 V=7.0 ACC=20 DEC=20
MOVL C00197 V=7.0 ACC=20 DEC=20
MOVL C00198 V=7.0 ACC=20 DEC=20
MOVL C00199 V=7.0 ACC=20 DEC=20
MOVL C00200 V=7.0 ACC=20 DEC=20
MOVL C00201 V=7.0 ACC=20 DEC=20
ARCOF
TIMER T=30
*LAG9
MOVL C00202 V=11.0 ACC=20 DEC=20
MACRO1 MJ#(0) ARGF2
ARCON
MOVL C00203 V=7.0 ACC=20 DEC=20
MOVL C00204 V=7.0 ACC=20 DEC=20
MOVL C00205 V=7.0 ACC=20 DEC=20
MOVL C00206 V=7.0 ACC=20 DEC=20
MOVL C00207 V=7.0 ACC=20 DEC=20
MOVL C00208 V=7.0 ACC=20 DEC=20
MOVL C00209 V=7.0 ACC=20 DEC=20
MOVL C00210 V=7.0 ACC=20 DEC=20
MOVL C00211 V=7.0 ACC=20 DEC=20
MOVL C00212 V=7.0 ACC=20 DEC=20
MOVL C00213 V=7.0 ACC=20 DEC=20
MOVL C00214 V=7.0 ACC=20 DEC=20
MOVL C00215 V=7.0 ACC=20 DEC=20
MOVL C00216 V=7.0 ACC=20 DEC=20
MOVL C00217 V=7.0 ACC=20 DEC=20
MOVL C00218 V=7.0 ACC=20 DEC=20
MOVL C00219 V=7.0 ACC=20 DEC=20
MOVL C00220 V=7.0 ACC=20 DEC=20
MOVL C00221 V=7.0 ACC=20 DEC=20
MOVL C00222 V=7.0 ACC=20 DEC=20
MOVL C00223 V=7.0 ACC=20 DEC=20
MOVL C00224 V=7.0 ACC=20 DEC=20
MOVL C00225 V=7.0 ACC=20 DEC=20
MOVL C00226 V=7.0 ACC=20 DEC=20
ARCOF
TIMER T=30
*LAG10
MOVL C00227 V=11.0 ACC=20 DEC=20
MACRO1 MJ#(0) ARGF2
ARCON
MOVL C00228 V=7.0 ACC=20 DEC=20
MOVL C00229 V=7.0 ACC=20 DEC=20
MOVL C00230 V=7.0 ACC=20 DEC=20
MOVL C00231 V=7.0 ACC=20 DEC=20
MOVL C00232 V=7.0 ACC=20 DEC=20
MOVL C00233 V=7.0 ACC=20 DEC=20
MOVL C00234 V=7.0 ACC=20 DEC=20
MOVL C00235 V=7.0 ACC=20 DEC=20
MOVL C00236 V=7.0 ACC=20 DEC=20
MOVL C00237 V=7.0 ACC=20 DEC=20
MOVL C00238 V=7.0 ACC=20 DEC=20
MOVL C00239 V=7.0 ACC=20 DEC=20
MOVL C00240 V=7.0 ACC=20 DEC=20
MOVL C00241 V=7.0 ACC=20 DEC=20
MOVL C00242 V=7.0 ACC=20 DEC=20
MOVL C00243 V=7.0 ACC=20 DEC=20
MOVL C00244 V=7.0 ACC=20 DEC=20
MOVL C00245 V=7.0 ACC=20 DEC=20
MOVL C00246 V=7.0 ACC=20 DEC=20
MOVL C00247 V=7.0 ACC=20 DEC=20
MOVL C00248 V=7.0 ACC=20 DEC=20
MOVL C00249 V=7.0 ACC=20 DEC=20
MOVL C00250 V=7.0 ACC=20 DEC=20
MOVL C00251 V=7.0 ACC=20 DEC=20
ARCOF
TIMER T=30
*LAG11
MOVL C00252 V=11.0 ACC=20 DEC=20
MACRO1 MJ#(0) ARGF2
ARCON
MOVL C00253 V=7.0 ACC=20 DEC=20
MOVL C00254 V=7.0 ACC=20 DEC=20
MOVL C00255 V=7.0 ACC=20 DEC=20
MOVL C00256 V=7.0 ACC=20 DEC=20
MOVL C00257 V=7.0 ACC=20 DEC=20
MOVL C00258 V=7.0 ACC=20 DEC=20
MOVL C00259 V=7.0 ACC=20 DEC=20
MOVL C00260 V=7.0 ACC=20 DEC=20
MOVL C00261 V=7.0 ACC=20 DEC=20
MOVL C00262 V=7.0 ACC=20 DEC=20
MOVL C00263 V=7.0 ACC=20 DEC=20
MOVL C00264 V=7.0 ACC=20 DEC=20
MOVL C00265 V=7.0 ACC=20 DEC=20
MOVL C00266 V=7.0 ACC=20 DEC=20
MOVL C00267 V=7.0 ACC=20 DEC=20
MOVL C00268 V=7.0 ACC=20 DEC=20
MOVL C00269 V=7.0 ACC=20 DEC=20
MOVL C00270 V=7.0 ACC=20 DEC=20
MOVL C00271 V=7.0 ACC=20 DEC=20
MOVL C00272 V=7.0 ACC=20 DEC=20
MOVL C00273 V=7.0 ACC=20 DEC=20
MOVL C00274 V=7.0 ACC=20 DEC=20
MOVL C00275 V=7.0 ACC=20 DEC=20
MOVL C00276 V=7.0 ACC=20 DEC=20
ARCOF
TIMER T=30
*LAG12
MOVL C00277 V=11.0 ACC=20 DEC=20
MACRO1 MJ#(0) ARGF2
ARCON
MOVL C00278 V=7.0 ACC=20 DEC=20
MOVL C00279 V=7.0 ACC=20 DEC=20
MOVL C00280 V=7.0 ACC=20 DEC=20
MOVL C00281 V=7.0 ACC=20 DEC=20
MOVL C00282 V=7.0 ACC=20 DEC=20
MOVL C00283 V=7.0 ACC=20 DEC=20
MOVL C00284 V=7.0 ACC=20 DEC=20
MOVL C00285 V=7.0 ACC=20 DEC=20
MOVL C00286 V=7.0 ACC=20 DEC=20
MOVL C00287 V=7.0 ACC=20 DEC=20
MOVL C00288 V=7.0 ACC=20 DEC=20
MOVL C00289 V=7.0 ACC=20 DEC=20
MOVL C00290 V=7.0 ACC=20 DEC=20
MOVL C00291 V=7.0 ACC=20 DEC=20
MOVL C00292 V=7.0 ACC=20 DEC=20
MOVL C00293 V=7.0 ACC=20 DEC=20
MOVL C00294 V=7.0 ACC=20 DEC=20
MOVL C00295 V=7.0 ACC=20 DEC=20
MOVL C00296 V=7.0 ACC=20 DEC=20
MOVL C00297 V=7.0 ACC=20 DEC=20
MOVL C00298 V=7.0 ACC=20 DEC=20
MOVL C00299 V=7.0 ACC=20 DEC=20
MOVL C00300 V=7.0 ACC=20 DEC=20
MOVL C00301 V=7.0 ACC=20 DEC=20
ARCOF
TIMER T=30
*LAG13
MOVL C00302 V=11.0 ACC=20 DEC=20
MACRO1 MJ#(0) ARGF2
ARCON
MOVL C00303 V=7.0 ACC=20 DEC=20
MOVL C00304 V=7.0 ACC=20 DEC=20
MOVL C00305 V=7.0 ACC=20 DEC=20
MOVL C00306 V=7.0 ACC=20 DEC=20
MOVL C00307 V=7.0 ACC=20 DEC=20
MOVL C00308 V=7.0 ACC=20 DEC=20
MOVL C00309 V=7.0 ACC=20 DEC=20
MOVL C00310 V=7.0 ACC=20 DEC=20
MOVL C00311 V=7.0 ACC=20 DEC=20
MOVL C00312 V=7.0 ACC=20 DEC=20
MOVL C00313 V=7.0 ACC=20 DEC=20
MOVL C00314 V=7.0 ACC=20 DEC=20
MOVL C00315 V=7.0 ACC=20 DEC=20
MOVL C00316 V=7.0 ACC=20 DEC=20
MOVL C00317 V=7.0 ACC=20 DEC=20
MOVL C00318 V=7.0 ACC=20 DEC=20
MOVL C00319 V=7.0 ACC=20 DEC=20
MOVL C00320 V=7.0 ACC=20 DEC=20
MOVL C00321 V=7.0 ACC=20 DEC=20
MOVL C00322 V=7.0 ACC=20 DEC=20
MOVL C00323 V=7.0 ACC=20 DEC=20
MOVL C00324 V=7.0 ACC=20 DEC=20
MOVL C00325 V=7.0 ACC=20 DEC=20
MOVL C00326 V=7.0 ACC=20 DEC=20
ARCOF
TIMER T=30
*LAG14
MOVL C00327 V=11.0 ACC=20 DEC=20
MACRO1 MJ#(0) ARGF2
ARCON
MOVL C00328 V=7.0 ACC=20 DEC=20
MOVL C00329 V=7.0 ACC=20 DEC=20
MOVL C00330 V=7.0 ACC=20 DEC=20
MOVL C00331 V=7.0 ACC=20 DEC=20
MOVL C00332 V=7.0 ACC=20 DEC=20
MOVL C00333 V=7.0 ACC=20 DEC=20
MOVL C00334 V=7.0 ACC=20 DEC=20
MOVL C00335 V=7.0 ACC=20 DEC=20
MOVL C00336 V=7.0 ACC=20 DEC=20
MOVL C00337 V=7.0 ACC=20 DEC=20
MOVL C00338 V=7.0 ACC=20 DEC=20
MOVL C00339 V=7.0 ACC=20 DEC=20
MOVL C00340 V=7.0 ACC=20 DEC=20
MOVL C00341 V=7.0 ACC=20 DEC=20
MOVL C00342 V=7.0 ACC=20 DEC=20
MOVL C00343 V=7.0 ACC=20 DEC=20
MOVL C00344 V=7.0 ACC=20 DEC=20
MOVL C00345 V=7.0 ACC=20 DEC=20
MOVL C00346 V=7.0 ACC=20 DEC=20
MOVL C00347 V=7.0 ACC=20 DEC=20
MOVL C00348 V=7.0 ACC=20 DEC=20
MOVL C00349 V=7.0 ACC=20 DEC=20
MOVL C00350 V=7.0 ACC=20 DEC=20
MOVL C00351 V=7.0 ACC=20 DEC=20
ARCOF
TIMER T=30
*LAG15
MOVL C00352 V=11.0 ACC=20 DEC=20
MACRO1 MJ#(0) ARGF2
ARCON
MOVL C00353 V=7.0 ACC=20 DEC=20
MOVL C00354 V=7.0 ACC=20 DEC=20
MOVL C00355 V=7.0 ACC=20 DEC=20
MOVL C00356 V=7.0 ACC=20 DEC=20
MOVL C00357 V=7.0 ACC=20 DEC=20
MOVL C00358 V=7.0 ACC=20 DEC=20
MOVL C00359 V=7.0 ACC=20 DEC=20
MOVL C00360 V=7.0 ACC=20 DEC=20
MOVL C00361 V=7.0 ACC=20 DEC=20
MOVL C00362 V=7.0 ACC=20 DEC=20
MOVL C00363 V=7.0 ACC=20 DEC=20
MOVL C00364 V=7.0 ACC=20 DEC=20
MOVL C00365 V=7.0 ACC=20 DEC=20
MOVL C00366 V=7.0 ACC=20 DEC=20
MOVL C00367 V=7.0 ACC=20 DEC=20
MOVL C00368 V=7.0 ACC=20 DEC=20
MOVL C00369 V=7.0 ACC=20 DEC=20
MOVL C00370 V=7.0 ACC=20 DEC=20
MOVL C00371 V=7.0 ACC=20 DEC=20
MOVL C00372 V=7.0 ACC=20 DEC=20
MOVL C00373 V=7.0 ACC=20 DEC=20
MOVL C00374 V=7.0 ACC=20 DEC=20
MOVL C00375 V=7.0 ACC=20 DEC=20
MOVL C00376 V=7.0 ACC=20 DEC=20
ARCOF
TIMER T=30
MOVL C00377 V=11.0 ACC=20 DEC=20
MOVJ C00378 VJ=0.78
END
